(* IEC 61131-3 sources: PortalRobot/Portal_robot/Device/application/ST/ST_POINT, 2 files *)

(* ---- E_POINT_NAME.st ---- *)
{attribute 'qualified_only'}
{attribute 'strict'}
TYPE E_POINT_NAME :
(
	NONE,
	MACHINE_1_ABOVE,
	MACHINE_1_INSIDE, // Legacy: исключена из редактора, сохранена ради числового протокола
	MACHINE_1_CHUCK_APROACH,
	MACHINE_1_CHUCK_POSITION,
	MACHINE_2_ABOVE,
	MACHINE_2_INSIDE, // Legacy: исключена из редактора, сохранена ради числового протокола
	MACHINE_2_CHUCK_APROACH,
	MACHINE_2_CHUCK_POSITION,
	MACHINE_3_ABOVE,
	MACHINE_3_INSIDE, // Legacy: исключена из редактора, сохранена ради числового протокола
	MACHINE_3_CHUCK_APROACH,
	MACHINE_3_CHUCK_POSITION,
	MAGAZINE_DETAIL,
	MAGAZINE_TAKE_DETAIL,
	MAGAZINE_PUT_DETAIL,
	MAGAZINE_CHANGE_DETAIL,
	HOME_SAFETY,
	MAGAZINE_RETURN_BLANK, // Legacy: сохранено только ради прежнего числового значения
	MAGAZINE_SAFE, // Безопасная точка над активным слотом
	MAGAZINE_IN_SLOT, // Рабочая точка внутри активного слота
	MAGAZINE_CHANGE, // Безопасная точка переворота над активным слотом
	MAGAZINE_1_DETAIL, // Базовая точка рабочей зоны первого магазина
	MAGAZINE_2_DETAIL, // Базовая точка рабочей зоны второго магазина
	GEOMETRY_1_PLACE,
	GEOMETRY_1_SAFE,
	GEOMETRY_1_CHANGE,
	GEOMETRY_2_PLACE,
	GEOMETRY_2_SAFE,
	GEOMETRY_2_CHANGE,
	MAGAZINE_1_AXIS_X, // B: последний слот первого ряда магазина 1
	MAGAZINE_1_AXIS_Y, // C: первый слот последнего ряда магазина 1
	MAGAZINE_2_AXIS_X,
	MAGAZINE_2_AXIS_Y

);
END_TYPE

(* ---- ST_POINT.st ---- *)
TYPE ST_POINT :
STRUCT
	Name        : STRING[80]; // Имя точки
	X           : LREAL; // Координата X
	Y           : LREAL; // Координата Y
	Z           : LREAL; // Координата Z
	MagazineSafeZ : LREAL; // Signed-смещение Safe Z базы магазина или ГК
	MagazineChangeZ : LREAL; // Signed-смещение Change Z; используется только базовой точкой магазина
	SpeedFactor : LREAL; // Коэффициент скорости движения
	xConfigured : BOOL; // Для базы магазина TRUE только при ненулевых MagazineSafeZ и MagazineChangeZ
END_STRUCT
END_TYPE
